// TIA Portal V20 export
Screen "Pop-up_PRODDATA_CT_LEGEND_Popup"  330x456
  ScreenItem "Background" at 0,0 size 330x456  Type=HmiRectangle
  ScreenItem "Textfeld_Legende" at 1,1 size 328x25  Type=HmiTextBox
  ScreenItem "Textfeld_11" at 70,364 size 255x88  Type=HmiTextBox
  ScreenItem "Textfeld_8" at 10,412 size 55x30  Type=HmiTextBox
  ScreenItem "Textfeld_9" at 23,392 size 30x20  Type=HmiTextBox
  ScreenItem "Textfeld_13" at 10,364 size 55x30  Type=HmiTextBox
  ScreenItem "Textfeld_10" at 10,34 size 205x28  Type=HmiTextBox
  ScreenItem "Textfeld_12" at 10,101 size 205x25  Type=HmiTextBox
  ScreenItem "Textfeld_14" at 10,64 size 318x35  Type=HmiTextBox
  ScreenItem "Textfeld_15" at 10,127 size 318x40  Type=HmiTextBox
  ScreenItem "Textfeld_2" at 10,218 size 55x30  Type=HmiTextBox
  ScreenItem "Textfeld_3" at 70,218 size 255x74  Type=HmiTextBox
  ScreenItem "Textfeld_4" at 10,251 size 55x30  Type=HmiTextBox
  ScreenItem "Textfeld_5" at 10,292 size 55x30  Type=HmiTextBox
  ScreenItem "Textfeld_6" at 70,292 size 255x70  Type=HmiTextBox
  ScreenItem "Textfeld_7" at 10,324 size 55x30  Type=HmiTextBox
  ScreenItem "Text_IONoMeasure" at 10,169 size 100x25  Type=HmiTextBox
  ScreenItem "Text_IOMeasureRun" at 115,169 size 100x25  Type=HmiTextBox
  ScreenItem "Text_IOMeasureHold" at 220,169 size 100x25  Type=HmiTextBox
  ScreenItem "Text_NoMeasure" at 10,195 size 100x20  Type=HmiTextBox
  ScreenItem "Text_MeasureRun" at 115,195 size 100x20  Type=HmiTextBox
  ScreenItem "Text_MeasureHold" at 220,195 size 100x20  Type=HmiTextBox
  ScreenItem "Cancel Mode" at 239,1 size 90x60  Type=HmiButton
